FUNCTION_BLOCK SortingSafeSequence (* The shared complete Stop procedure used for Stop commands and operating faults. *)
  (* Standard: 61499-2 *)
  (* Version 2.0, 2026-11-09, sorting2n, sorting2n *)
  PACKAGE Main;
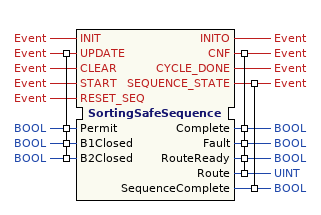
  EVENT_INPUT
    INIT;
    UPDATE WITH Permit, B1Closed, B2Closed;
    CLEAR;
    START;
    RESET_SEQ;
  END_EVENT
  EVENT_OUTPUT
    INITO;
    CNF WITH Complete, Fault, RouteReady, Route;
    CYCLE_DONE;
    SEQUENCE_STATE WITH SequenceComplete;
  END_EVENT
  VAR_INPUT
    Permit : BOOL := FALSE;
    B1Closed : BOOL;
    B2Closed : BOOL;
  END_VAR
  VAR_OUTPUT
    Complete : BOOL;
    Fault : BOOL;
    RouteReady : BOOL;
    Route : UINT := 0;
    SequenceComplete : BOOL;
  END_VAR
  FBS
    Flow : SortingSafeSteps; (* Standard safe-position sequence and its original timing. *)
    Services : SortingSafeServices; (* Existing ownership, command and measured home conditions. *)
  END_FBS
  EVENT_CONNECTIONS
    INIT TO Services.9406177C96964918;
    Flow.F1C83D723563445B TO CNF;
    UPDATE TO Services.B487FBD83E664405;
    Services.44AB9629DFF24FF7 TO INITO;
    UPDATE TO Flow.92A86B7AE0974DC0;
    Services.81C67910DE5D4FBE TO CNF;
    CLEAR TO Services.C03E480D6990400D;
    START TO Flow.378554B1BB2249B1;
    RESET_SEQ TO Flow.AC1D5F5E28444264;
    Flow.C7573A889A014538 TO SEQUENCE_STATE;
  END_CONNECTIONS
  DATA_CONNECTIONS
    Flow.44C30F2646B04FB5 TO Complete;
    B1Closed TO Services.39B88A85D9E443EC;
    B2Closed TO Services.819D37304DF54BE0;
    Services.33BD2F3DC21A43C2 TO Fault;
    Flow.A37666370B934C10 TO SequenceComplete;
  END_CONNECTIONS
  ADAPTER_CONNECTIONS
    Flow.132BF54BC9E64B19 TO Services.59D40A58A22B4030;
  END_CONNECTIONS
END_FUNCTION_BLOCK
